(* IEC 61131-3 sources: PLC-Static-Analysis/modules/plc-rules/src/test/resources/PLCA-L023, 2 files *)

(* ---- compliant.st ---- *)
FUNCTION F_L023ok : INT
VAR_INPUT
    nRaw : INT;
    b : BOOL;
END_VAR
VAR
    nTmp : INT;
    p : POINTER TO INT;
    nAlias : INT;
END_VAR
nTmp := nRaw * 2;
nTmp := nTmp + 1;
nTmp := nTmp * nRaw;
IF b THEN
    nTmp := 0;
END_IF
F_L023ok := nTmp;
p := ADR(nAlias);
nAlias := 1;
nAlias := 2;
nTmp := ABS(nRaw);
nTmp := 5;
F_L023ok := nTmp + p^;
END_FUNCTION

FUNCTION_BLOCK FB_L023ok
VAR_INPUT
    nRaw : INT;
END_VAR
VAR
    nStat : INT;
END_VAR
nStat := nRaw;
nStat := nRaw + 1;
END_FUNCTION_BLOCK

(* ---- noncompliant.st ---- *)
FUNCTION F_L023 : INT
VAR_INPUT
    nRaw : INT;
    b : BOOL;
END_VAR
VAR
    nTmp : INT;
    nOther : INT;
END_VAR
nTmp := nRaw * 2; // PLCA-L023
nTmp := nRaw * 3;
nOther := 1; // PLCA-L023
IF b THEN
    nTmp := 0;
END_IF
nOther := 2;
F_L023 := nTmp + nOther;
END_FUNCTION

FUNCTION_BLOCK FB_L023
VAR_INPUT
    nRaw : INT;
END_VAR
VAR_OUTPUT
    nOut : INT;
END_VAR
VAR_TEMP
    nTmp : INT;
END_VAR
nTmp := nRaw; // PLCA-L023
nTmp := nRaw + 1;
nOut := nTmp;
END_FUNCTION_BLOCK
